(* Logix 5000 project; controller R400_500_XLS vendor 1 type 14 code 216 rev 31.11; software revision 31.01; part 23 of 32 *)
(* tags used below, declared in another part *)
   Abort1 : DINT;   // Not Used
   Alarm : SINT;   // Wait 3 seconds
   AlarmAcked : BOOL;   // Alarm has been acked
   bAlrm : BOOL[64];
   CycExcBuffer : UDT_CYCLE;
   CycleSequence : UDT_CYCLE_SEQUENCE;
   DrnSmp : DINT;
   DRYING : DINT;   // Drying id number
   drying_sp : REAL;   // Drying temperature set point
   drying_sp_offset : REAL;   // Low drying offset
   DRYING_TEMP_HIGH : REAL;   // Smart drying high temperature set point
   DRYING_TEMP_LOW : REAL;   // Smart drying low temperature set point
   DRYING_TEMP_STANDARD_LOW : REAL;   // Regular drying low temperature set point
   DRYING_TIME_LONG : DINT;   // Smart drying time for heat sensitive mode (in minute)
   DRYING_TIME_SHORT : DINT;   // Smart drying time for heat regular mode (in minute)
   dryingSmartTime : DINT;   // Duration of the smart drying phase
   DryingTempCool : REAL;   // Temperature limit for the smart drying mode cooling phase
   F2rinse : DINT;   // Not Used
   F3rinse : DINT;   // Not Used
   F4rinse : INT;   // Transition for the conductivity based evalutaion
   F4rinse_Tran : INT;   // Transitions for the conductivity based evaluation
   Fill_Sump : DINT;
   FRinseCondValue : REAL;   // Stored value of the conductivity
   HeatSmp : DINT;
   Inj_Time : SINT;   // Time based chemical injection steps
   M : DINT[5];   // Memory Bits
   NbFinalRinseDone : DINT;
   Neutral : SINT;
   ONS_FC08 : DINT;
   ONS_FC09 : SINT;
   PureWaterTankFilling : BOOL;   // Start PWT filling
   Run : DINT;
   STANDARD : SINT;
   SumpWaterVolume : DINT;   // Sump Water Volume 0 =Low 1= High
   Tmr : TIMER[107];
   Treatment_info : DINT;   // Treatment message conditions
   Trt_Drying : SINT;
   Trt_Drying_Tran : INT;
   Trt_Vapor_Exhaust : BOOL;   // Vapor exhaust fan is on
   VENTING : DINT;   // Venting id number
   WaterSaved : BOOL;   // Water Saved In Sump (Last Final Rinse Water)
   WSH56_TreatmentInfo : BOOL;   // Treatment information for the conductivity injection
   COOLING_PHASE_TIME : DINT;   // Time of the cooling phase when time based drying
   DryTemp : REAL;
   FALSE : BOOL;   // Always false bit
   FinalRinseCond : REAL;
   Msg_Phase : DINT;
   PrintFrinseCondValue : REAL;
   PureWaterTankDrainingDeadLeg : BOOL;
   PureWaterTankFillingRequest : BOOL;
   Q_Smp_Stm_Vlve : BOOL;   // Sump steam valve/ Electrical Heater
   TreatmentPtr : DINT;
   Unit : Hrdwre;   // Unit Configuration
(* MainProgram, continued *)

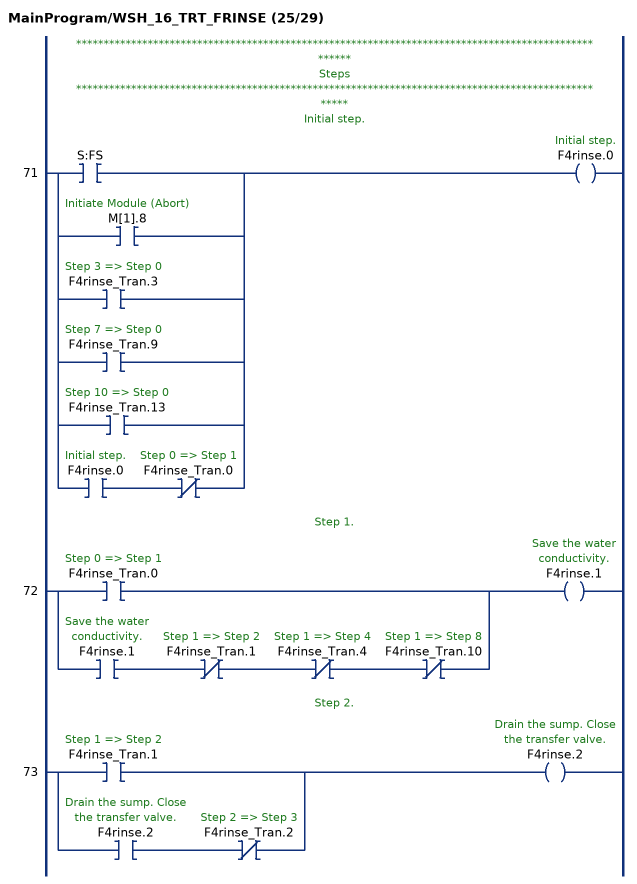
   [picture p449: MainProgram/WSH_16_TRT_FRINSE rungs 71-73]
   // ****************************************************************************************************
   // Steps
   // ***************************************************************************************************
   // Initial step.
   71: [XIC(S:FS) ,XIC(M[1].8) ,XIC(F4rinse_Tran.3) ,XIC(F4rinse_Tran.9) ,XIC(F4rinse_Tran.13) ,XIC(F4rinse.0) XIO(F4rinse_Tran.0) ]OTE(F4rinse.0);
   // Step 1.
   72: [XIC(F4rinse_Tran.0) ,XIC(F4rinse.1) XIO(F4rinse_Tran.1) XIO(F4rinse_Tran.4) XIO(F4rinse_Tran.10) ]OTE(F4rinse.1);
   // Step 2.
   73: [XIC(F4rinse_Tran.1) ,XIC(F4rinse.2) XIO(F4rinse_Tran.2) ]OTE(F4rinse.2);
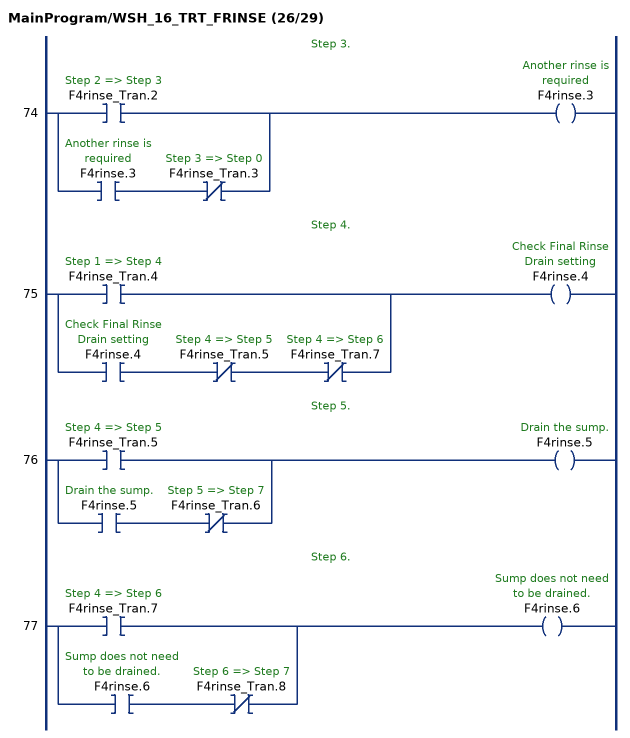
   // Step 3.
   74: [XIC(F4rinse_Tran.2) ,XIC(F4rinse.3) XIO(F4rinse_Tran.3) ]OTE(F4rinse.3);
   // Step 4.
   75: [XIC(F4rinse_Tran.4) ,XIC(F4rinse.4) XIO(F4rinse_Tran.5) XIO(F4rinse_Tran.7) ]OTE(F4rinse.4);
   // Step 5.
   76: [XIC(F4rinse_Tran.5) ,XIC(F4rinse.5) XIO(F4rinse_Tran.6) ]OTE(F4rinse.5);
   // Step 6.
   77: [XIC(F4rinse_Tran.7) ,XIC(F4rinse.6) XIO(F4rinse_Tran.8) ]OTE(F4rinse.6);
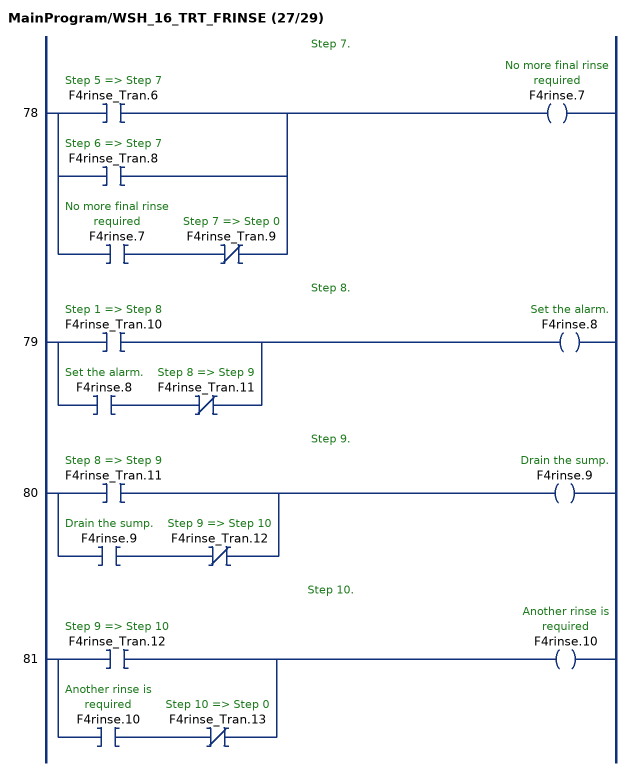
   // Step 7.
   78: [XIC(F4rinse_Tran.6) ,XIC(F4rinse_Tran.8) ,XIC(F4rinse.7) XIO(F4rinse_Tran.9) ]OTE(F4rinse.7);
   // Step 8.
   79: [XIC(F4rinse_Tran.10) ,XIC(F4rinse.8) XIO(F4rinse_Tran.11) ]OTE(F4rinse.8);
   // Step 9.
   80: [XIC(F4rinse_Tran.11) ,XIC(F4rinse.9) XIO(F4rinse_Tran.12) ]OTE(F4rinse.9);
   // Step 10.
   81: [XIC(F4rinse_Tran.12) ,XIC(F4rinse.10) XIO(F4rinse_Tran.13) ]OTE(F4rinse.10);
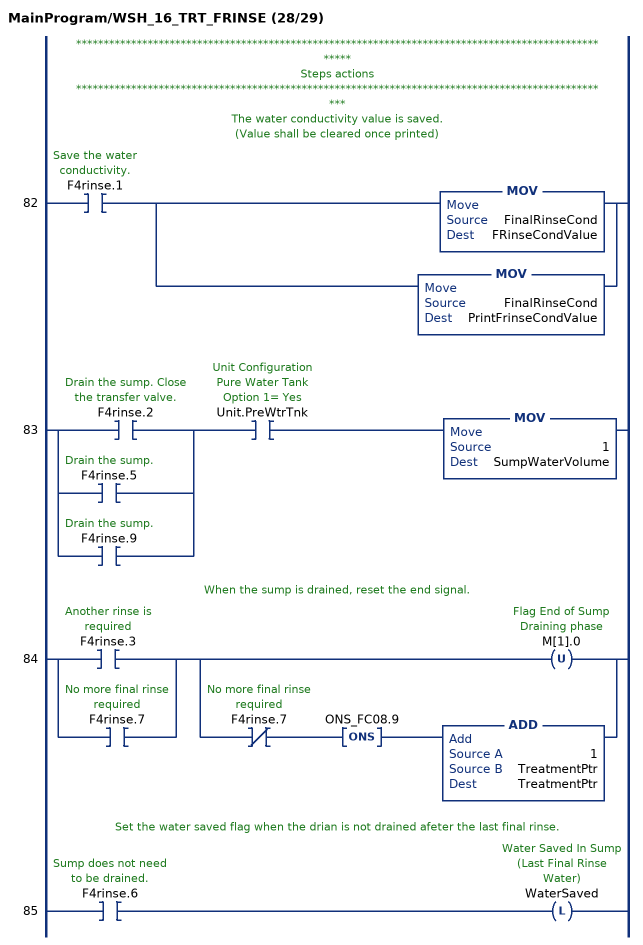
   // ****************************************************************************************************
   // Steps actions
   // **************************************************************************************************
   // The water conductivity value is saved.
   // (Value shall be cleared once printed)
   82: XIC(F4rinse.1)[MOV(FinalRinseCond,FRinseCondValue) ,MOV(FinalRinseCond,PrintFrinseCondValue) ];
   83: [XIC(F4rinse.2) ,XIC(F4rinse.5) ,XIC(F4rinse.9) ]XIC(Unit.PreWtrTnk)MOV(1,SumpWaterVolume);
   // When the sump is drained, reset the end signal.
   84: [XIC(F4rinse.3) ,XIC(F4rinse.7) ][OTU(M[1].0) ,XIO(F4rinse.7) ONS(ONS_FC08.9) ADD(1,TreatmentPtr,TreatmentPtr) ];
   // Set the water saved flag when the drian is not drained afeter the last final rinse.
   85: XIC(F4rinse.6)OTL(WaterSaved);
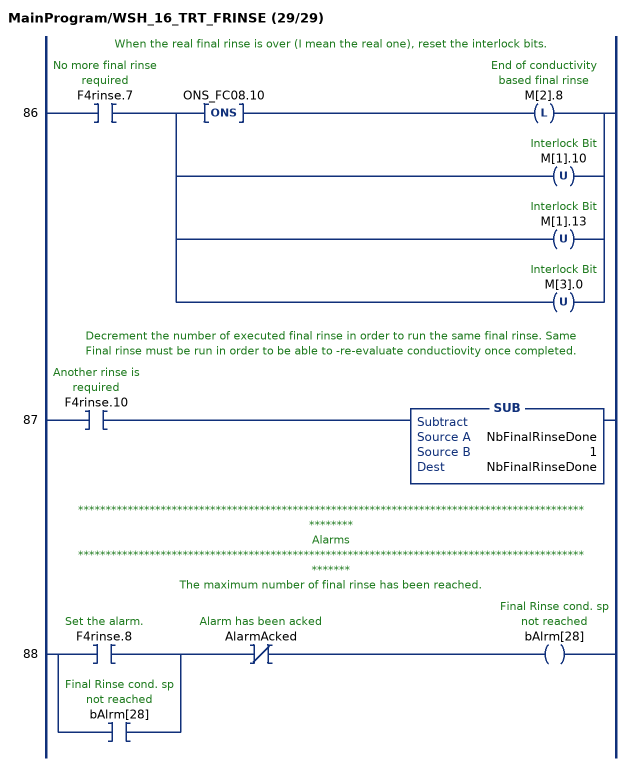
   // When the real final rinse is over (I mean the real one), reset the interlock bits.
   86: XIC(F4rinse.7)[ONS(ONS_FC08.10) OTL(M[2].8) ,OTU(M[1].10) ,OTU(M[1].13) ,OTU(M[3].0) ];
   // Decrement the number of executed final rinse in order to run the same final rinse. Same Final rinse must be run in order to be able to -re-evaluate conductiovity once completed.
   87: XIC(F4rinse.10)SUB(NbFinalRinseDone,1,NbFinalRinseDone);
   // ****************************************************************************************************
   // Alarms
   // ***************************************************************************************************
   // The maximum number of final rinse has been reached.
   88: [XIC(F4rinse.8) ,XIC(bAlrm[28]) ]XIO(AlarmAcked)OTE(bAlrm[28]);
END_ROUTINE

ROUTINE WSH_18_DRYING   (* ladder *)
// ROUTINe
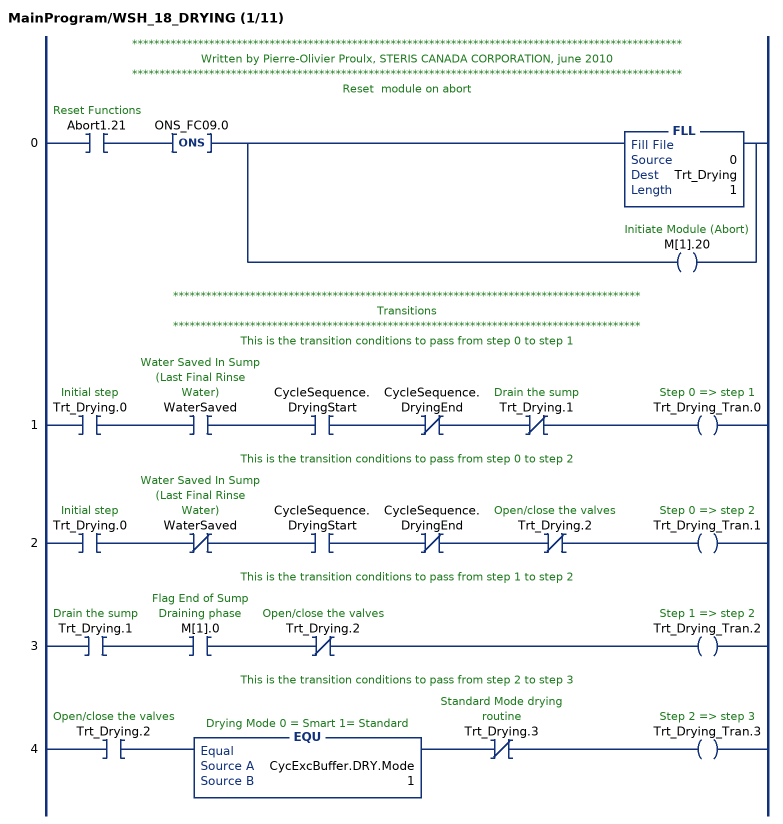
   // ****************************************************************************************************
   // Written by Pierre-Olivier Proulx, STERIS CANADA CORPORATION, june 2010
   // ****************************************************************************************************
   // Reset  module on abort
   0: XIC(Abort1.21)ONS(ONS_FC09.0)[FLL(0,Trt_Drying,1) ,OTE(M[1].20) ];
   // *************************************************************************************
   // Transitions
   // *************************************************************************************
   // This is the transition conditions to pass from step 0 to step 1
   1: XIC(Trt_Drying.0)XIC(WaterSaved)XIC(CycleSequence.DryingStart)XIO(CycleSequence.DryingEnd)XIO(Trt_Drying.1)OTE(Trt_Drying_Tran.0);
   // This is the transition conditions to pass from step 0 to step 2
   2: XIC(Trt_Drying.0)XIO(WaterSaved)XIC(CycleSequence.DryingStart)XIO(CycleSequence.DryingEnd)XIO(Trt_Drying.2)OTE(Trt_Drying_Tran.1);
   // This is the transition conditions to pass from step 1 to step 2
   3: XIC(Trt_Drying.1)XIC(M[1].0)XIO(Trt_Drying.2)OTE(Trt_Drying_Tran.2);
   // This is the transition conditions to pass from step 2 to step 3
   4: XIC(Trt_Drying.2)EQU(CycExcBuffer.DRY.Mode,1)XIO(Trt_Drying.3)OTE(Trt_Drying_Tran.3);
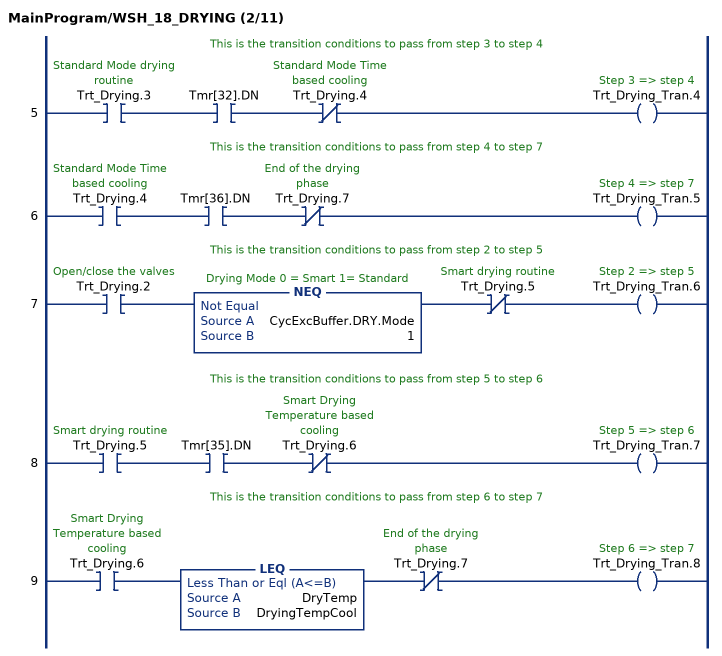
   // This is the transition conditions to pass from step 3 to step 4
   5: XIC(Trt_Drying.3)XIC(Tmr[32].DN)XIO(Trt_Drying.4)OTE(Trt_Drying_Tran.4);
   // This is the transition conditions to pass from step 4 to step 7
   6: XIC(Trt_Drying.4)XIC(Tmr[36].DN)XIO(Trt_Drying.7)OTE(Trt_Drying_Tran.5);
   // This is the transition conditions to pass from step 2 to step 5
   7: XIC(Trt_Drying.2)NEQ(CycExcBuffer.DRY.Mode,1)XIO(Trt_Drying.5)OTE(Trt_Drying_Tran.6);
   // This is the transition conditions to pass from step 5 to step 6
   8: XIC(Trt_Drying.5)XIC(Tmr[35].DN)XIO(Trt_Drying.6)OTE(Trt_Drying_Tran.7);
   // This is the transition conditions to pass from step 6 to step 7
   9: XIC(Trt_Drying.6)LEQ(DryTemp,DryingTempCool)XIO(Trt_Drying.7)OTE(Trt_Drying_Tran.8);
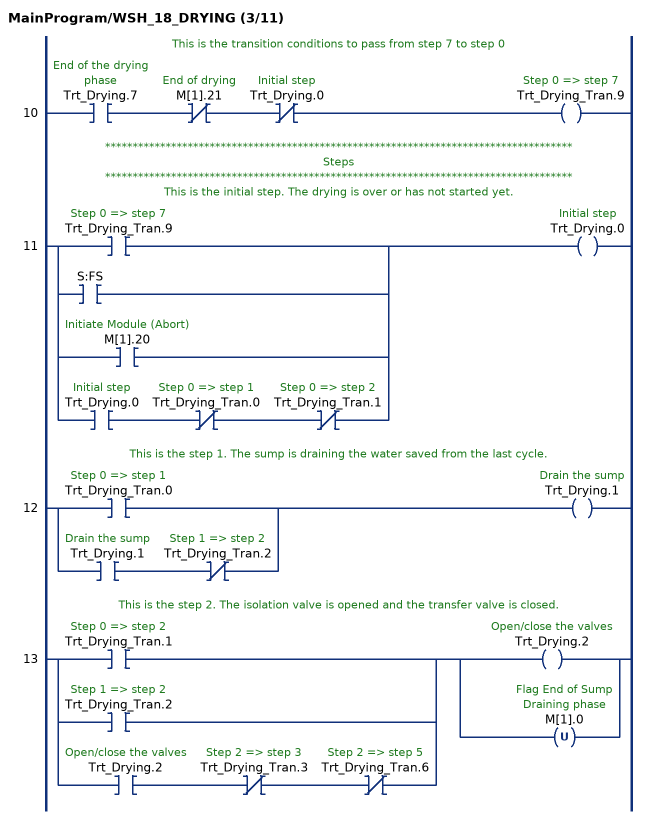
   // This is the transition conditions to pass from step 7 to step 0
   10: XIC(Trt_Drying.7)XIO(M[1].21)XIO(Trt_Drying.0)OTE(Trt_Drying_Tran.9);
   // *************************************************************************************
   // Steps
   // *************************************************************************************
   // This is the initial step. The drying is over or has not started yet.
   11: [XIC(Trt_Drying_Tran.9) ,XIC(S:FS) ,XIC(M[1].20) ,XIC(Trt_Drying.0) XIO(Trt_Drying_Tran.0) XIO(Trt_Drying_Tran.1) ]OTE(Trt_Drying.0);
   // This is the step 1. The sump is draining the water saved from the last cycle.
   12: [XIC(Trt_Drying_Tran.0) ,XIC(Trt_Drying.1) XIO(Trt_Drying_Tran.2) ]OTE(Trt_Drying.1);
   // This is the step 2. The isolation valve is opened and the transfer valve is closed.
   13: [XIC(Trt_Drying_Tran.1) ,XIC(Trt_Drying_Tran.2) ,XIC(Trt_Drying.2) XIO(Trt_Drying_Tran.3) XIO(Trt_Drying_Tran.6) ][OTE(Trt_Drying.2) ,OTU(M[1].0) ];
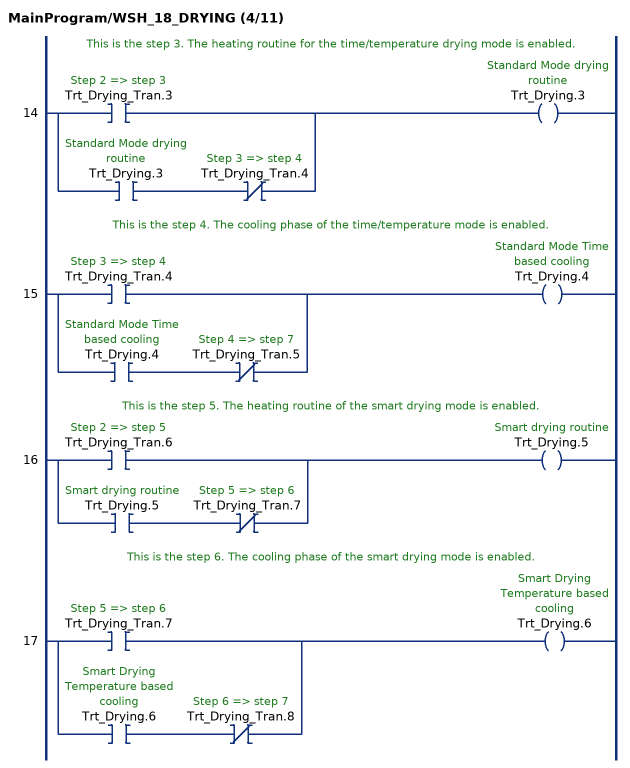
   // This is the step 3. The heating routine for the time/temperature drying mode is enabled.
   14: [XIC(Trt_Drying_Tran.3) ,XIC(Trt_Drying.3) XIO(Trt_Drying_Tran.4) ]OTE(Trt_Drying.3);
   // This is the step 4. The cooling phase of the time/temperature mode is enabled.
   15: [XIC(Trt_Drying_Tran.4) ,XIC(Trt_Drying.4) XIO(Trt_Drying_Tran.5) ]OTE(Trt_Drying.4);
   // This is the step 5. The heating routine of the smart drying mode is enabled.
   16: [XIC(Trt_Drying_Tran.6) ,XIC(Trt_Drying.5) XIO(Trt_Drying_Tran.7) ]OTE(Trt_Drying.5);
   // This is the step 6. The cooling phase of the smart drying mode is enabled.
   17: [XIC(Trt_Drying_Tran.7) ,XIC(Trt_Drying.6) XIO(Trt_Drying_Tran.8) ]OTE(Trt_Drying.6);
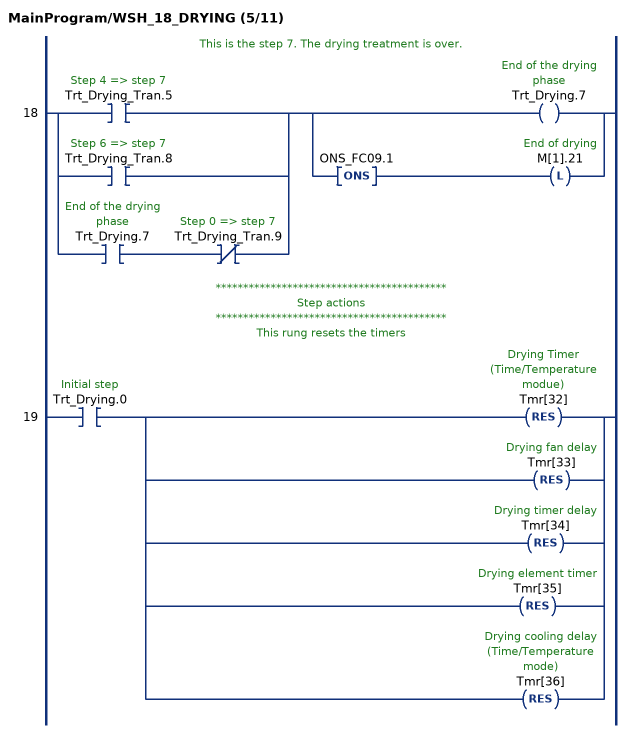
   // This is the step 7. The drying treatment is over.
   18: [XIC(Trt_Drying_Tran.5) ,XIC(Trt_Drying_Tran.8) ,XIC(Trt_Drying.7) XIO(Trt_Drying_Tran.9) ][OTE(Trt_Drying.7) ,ONS(ONS_FC09.1) OTL(M[1].21) ];
   // ******************************************
   // Step actions
   // ******************************************
   // This rung resets the timers
   19: XIC(Trt_Drying.0)[RES(Tmr[32]) ,RES(Tmr[33]) ,RES(Tmr[34]) ,RES(Tmr[35]) ,RES(Tmr[36]) ];
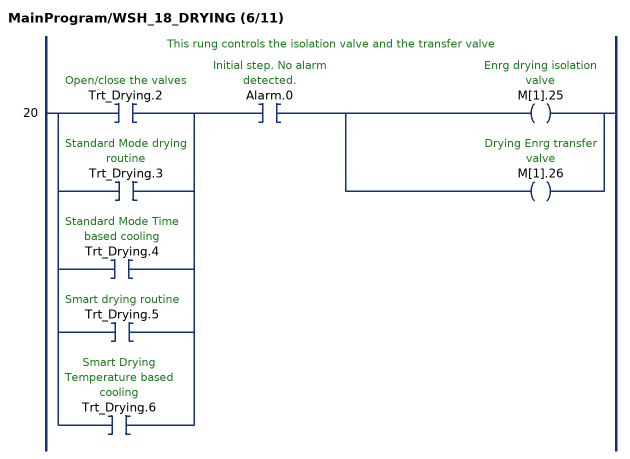
   // This rung controls the isolation valve and the transfer valve
   20: [XIC(Trt_Drying.2) ,XIC(Trt_Drying.3) ,XIC(Trt_Drying.4) ,XIC(Trt_Drying.5) ,XIC(Trt_Drying.6) ]XIC(Alarm.0)[OTE(M[1].25) ,OTE(M[1].26) ];
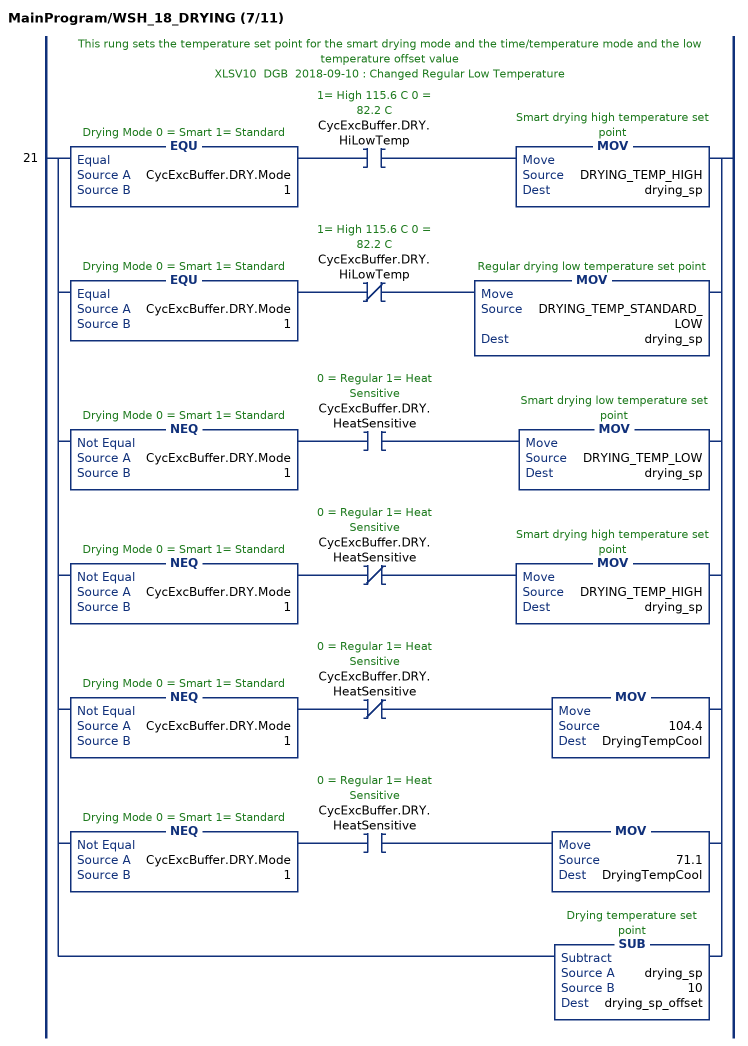
   // This rung sets the temperature set point for the smart drying mode and the time/temperature mode and the low temperature offset value
   // XLSV10  DGB  2018-09-10 : Changed Regular Low Temperature
   21: [EQU(CycExcBuffer.DRY.Mode,1) XIC(CycExcBuffer.DRY.HiLowTemp) MOV(DRYING_TEMP_HIGH,drying_sp) ,EQU(CycExcBuffer.DRY.Mode,1) XIO(CycExcBuffer.DRY.HiLowTemp) MOV(DRYING_TEMP_STANDARD_LOW,drying_sp) ,NEQ(CycExcBuffer.DRY.Mode,1) XIC(CycExcBuffer.DRY.HeatSensitive) MOV(DRYING_TEMP_LOW,drying_sp) ,NEQ(CycExcBuffer.DRY.Mode,1) XIO(CycExcBuffer.DRY.HeatSensitive) MOV(DRYING_TEMP_HIGH,drying_sp) ,NEQ(CycExcBuffer.DRY.Mode,1) XIO(CycExcBuffer.DRY.HeatSensitive) MOV(104.4,DryingTempCool) ,NEQ(CycExcBuffer.DRY.Mode,1) XIC(CycExcBuffer.DRY.HeatSensitive) MOV(71.1,DryingTempCool) ,SUB(drying_sp,10,drying_sp_offset) ];
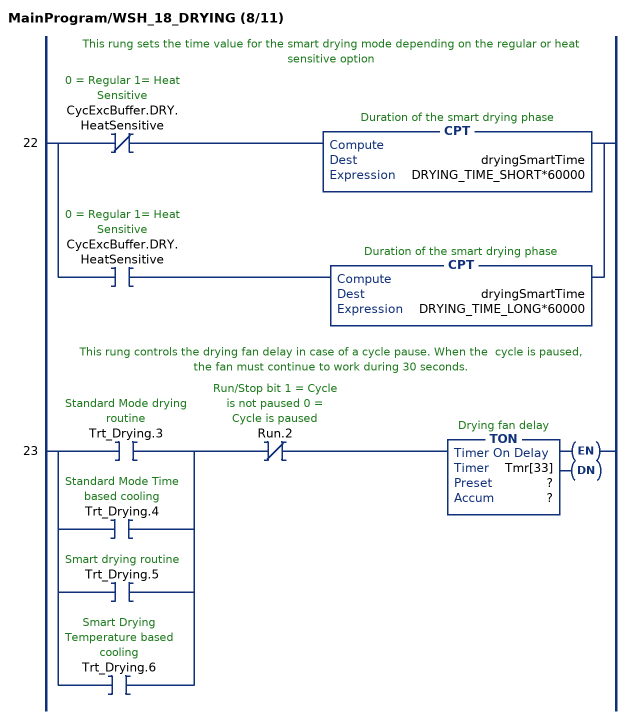
   // This rung sets the time value for the smart drying mode depending on the regular or heat sensitive option
   22: [XIO(CycExcBuffer.DRY.HeatSensitive) CPT(dryingSmartTime,DRYING_TIME_SHORT*60000) ,XIC(CycExcBuffer.DRY.HeatSensitive) CPT(dryingSmartTime,DRYING_TIME_LONG*60000) ];
   // This rung controls the drying fan delay in case of a cycle pause. When the  cycle is paused, the fan must continue to work during 30 seconds.
   23: [XIC(Trt_Drying.3) ,XIC(Trt_Drying.4) ,XIC(Trt_Drying.5) ,XIC(Trt_Drying.6) ]XIO(Run.2)TON(Tmr[33],?,?);
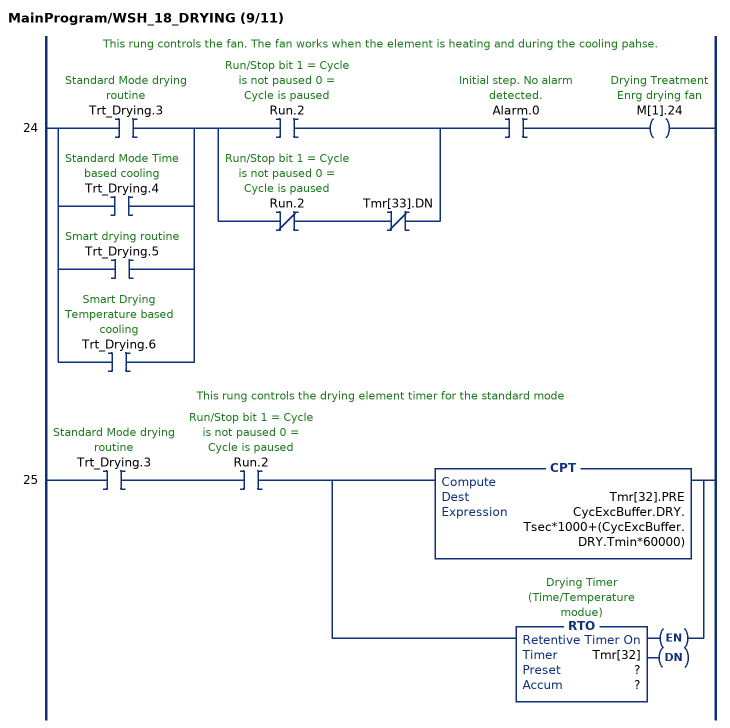
   // This rung controls the fan. The fan works when the element is heating and during the cooling pahse.
   24: [XIC(Trt_Drying.3) ,XIC(Trt_Drying.4) ,XIC(Trt_Drying.5) ,XIC(Trt_Drying.6) ][XIC(Run.2) ,XIO(Run.2) XIO(Tmr[33].DN) ]XIC(Alarm.0)OTE(M[1].24);
   // This rung controls the drying element timer for the standard mode
   25: XIC(Trt_Drying.3)XIC(Run.2)[CPT(Tmr[32].PRE,CycExcBuffer.DRY.Tsec*1000+(CycExcBuffer.DRY.Tmin*60000)) ,RTO(Tmr[32],?,?) ];
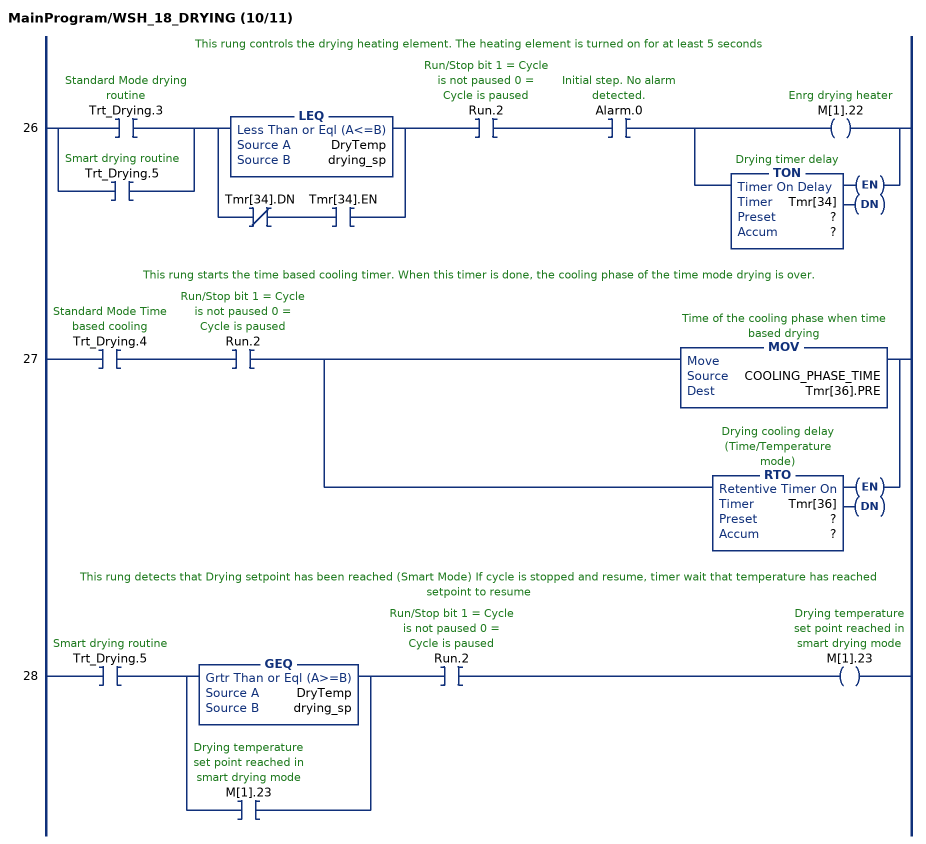
   // This rung controls the drying heating element. The heating element is turned on for at least 5 seconds
   26: [XIC(Trt_Drying.3) ,XIC(Trt_Drying.5) ][LEQ(DryTemp,drying_sp) ,XIO(Tmr[34].DN) XIC(Tmr[34].EN) ]XIC(Run.2)XIC(Alarm.0)[OTE(M[1].22) ,TON(Tmr[34],?,?) ];
   // This rung starts the time based cooling timer. When this timer is done, the cooling phase of the time mode drying is over.
   27: XIC(Trt_Drying.4)XIC(Run.2)[MOV(COOLING_PHASE_TIME,Tmr[36].PRE) ,RTO(Tmr[36],?,?) ];
   // This rung detects that Drying setpoint has been reached (Smart Mode) If cycle is stopped and resume, timer wait that temperature has reached setpoint to resume
   28: XIC(Trt_Drying.5)[GEQ(DryTemp,drying_sp) ,XIC(M[1].23) ]XIC(Run.2)OTE(M[1].23);
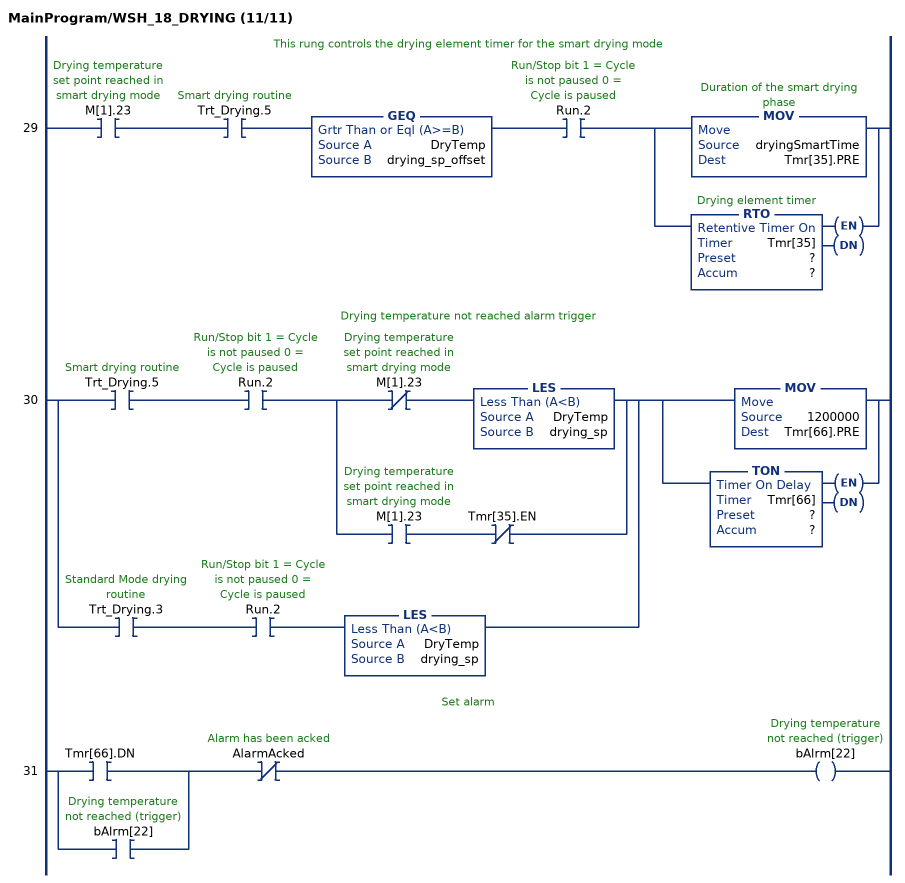
   // This rung controls the drying element timer for the smart drying mode
   29: XIC(M[1].23)XIC(Trt_Drying.5)GEQ(DryTemp,drying_sp_offset)XIC(Run.2)[MOV(dryingSmartTime,Tmr[35].PRE) ,RTO(Tmr[35],?,?) ];
   // Drying temperature not reached alarm trigger
   30: [XIC(Trt_Drying.5) XIC(Run.2) [XIO(M[1].23) LES(DryTemp,drying_sp) ,XIC(M[1].23) XIO(Tmr[35].EN) ] ,XIC(Trt_Drying.3) XIC(Run.2) LES(DryTemp,drying_sp) ][MOV(1200000,Tmr[66].PRE) ,TON(Tmr[66],?,?) ];
   // Set alarm
   31: [XIC(Tmr[66].DN) ,XIC(bAlrm[22]) ]XIO(AlarmAcked)OTE(bAlrm[22]);
END_ROUTINE

ROUTINE WSH_19_VENTING   (* ladder *)
// This routine vents the chamber
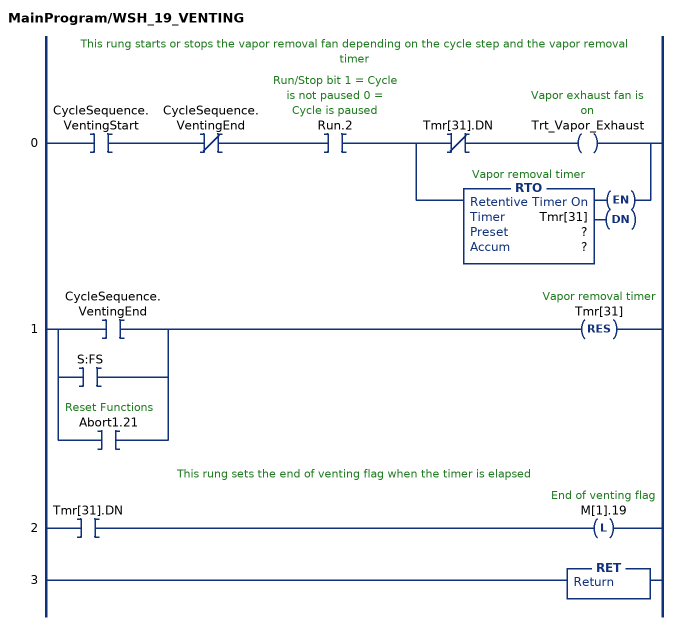
   // This rung starts or stops the vapor removal fan depending on the cycle step and the vapor removal timer
   0: XIC(CycleSequence.VentingStart)XIO(CycleSequence.VentingEnd)XIC(Run.2)[XIO(Tmr[31].DN) OTE(Trt_Vapor_Exhaust) ,RTO(Tmr[31],?,?) ];
   1: [XIC(CycleSequence.VentingEnd) ,[XIC(S:FS) ,XIC(Abort1.21) ] ]RES(Tmr[31]);
   // This rung sets the end of venting flag when the timer is elapsed
   2: XIC(Tmr[31].DN)OTL(M[1].19);
   3: RET();
END_ROUTINE

ROUTINE WSH_20_TREATMENT_INFO   (* ladder *)
// This routine decides which message the HMI will display during a cycle
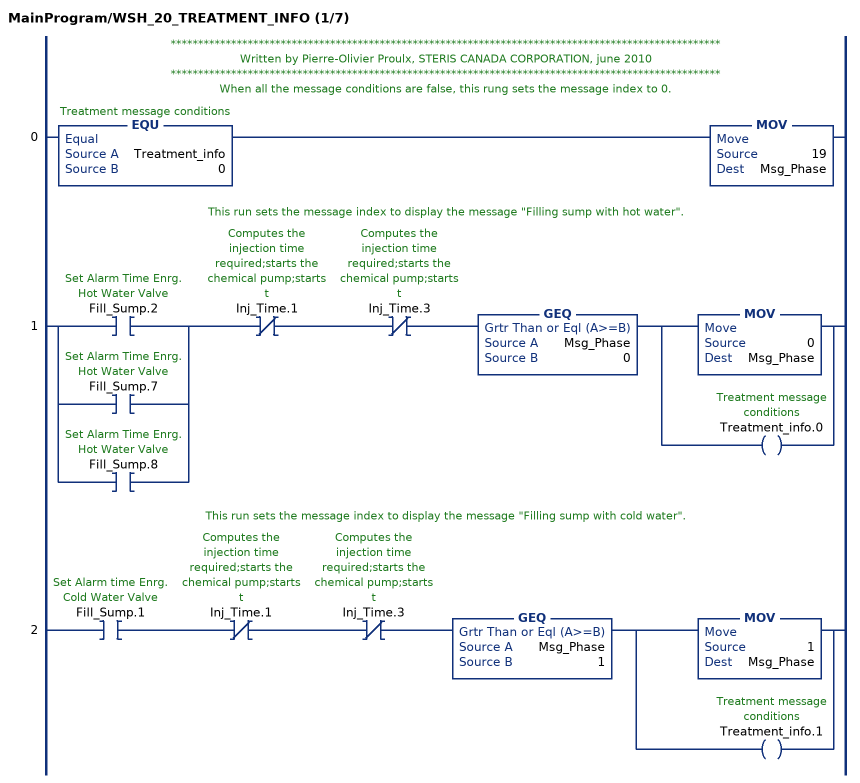
   // ****************************************************************************************************
   // Written by Pierre-Olivier Proulx, STERIS CANADA CORPORATION, june 2010
   // ****************************************************************************************************
   // When all the message conditions are false, this rung sets the message index to 0.
   0: EQU(Treatment_info,0)MOV(19,Msg_Phase);
   // This run sets the message index to display the message "Filling sump with hot water".
   1: [XIC(Fill_Sump.2) ,XIC(Fill_Sump.7) ,XIC(Fill_Sump.8) ]XIO(Inj_Time.1)XIO(Inj_Time.3)GEQ(Msg_Phase,0)[MOV(0,Msg_Phase) ,OTE(Treatment_info.0) ];
   // This run sets the message index to display the message "Filling sump with cold water".
   2: XIC(Fill_Sump.1)XIO(Inj_Time.1)XIO(Inj_Time.3)GEQ(Msg_Phase,1)[MOV(1,Msg_Phase) ,OTE(Treatment_info.1) ];
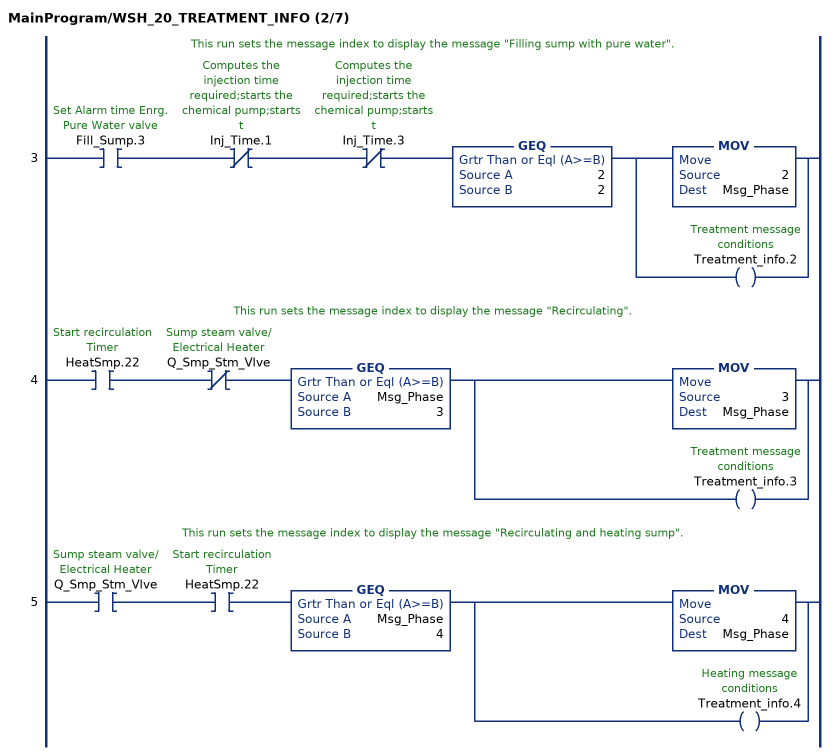
   // This run sets the message index to display the message "Filling sump with pure water".
   3: XIC(Fill_Sump.3)XIO(Inj_Time.1)XIO(Inj_Time.3)GEQ(2,2)[MOV(2,Msg_Phase) ,OTE(Treatment_info.2) ];
   // This run sets the message index to display the message "Recirculating".
   4: XIC(HeatSmp.22)XIO(Q_Smp_Stm_Vlve)GEQ(Msg_Phase,3)[MOV(3,Msg_Phase) ,OTE(Treatment_info.3) ];
   // This run sets the message index to display the message "Recirculating and heating sump".
   5: XIC(Q_Smp_Stm_Vlve)XIC(HeatSmp.22)GEQ(Msg_Phase,4)[MOV(4,Msg_Phase) ,OTE(Treatment_info.4) ];
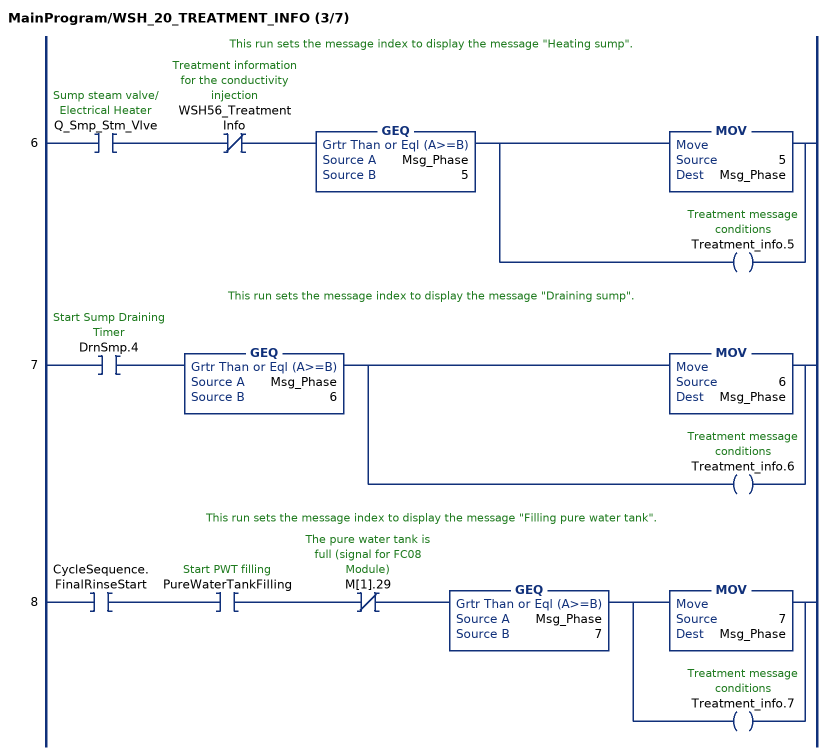
   // This run sets the message index to display the message "Heating sump".
   6: XIC(Q_Smp_Stm_Vlve)XIO(WSH56_TreatmentInfo)GEQ(Msg_Phase,5)[MOV(5,Msg_Phase) ,OTE(Treatment_info.5) ];
   // This run sets the message index to display the message "Draining sump".
   7: XIC(DrnSmp.4)GEQ(Msg_Phase,6)[MOV(6,Msg_Phase) ,OTE(Treatment_info.6) ];
   // This run sets the message index to display the message "Filling pure water tank".
   8: XIC(CycleSequence.FinalRinseStart)XIC(PureWaterTankFilling)XIO(M[1].29)GEQ(Msg_Phase,7)[MOV(7,Msg_Phase) ,OTE(Treatment_info.7) ];
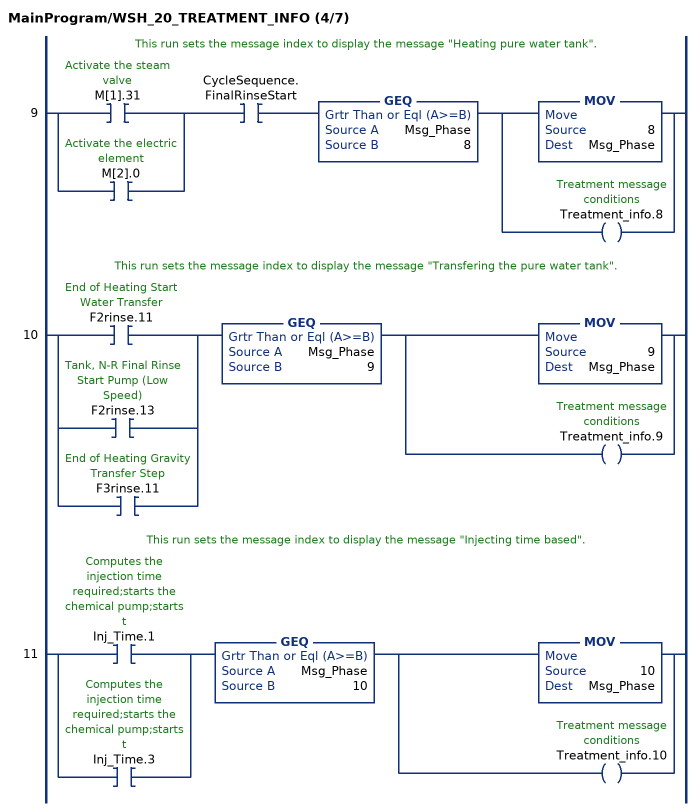
   // This run sets the message index to display the message "Heating pure water tank".
   9: [XIC(M[1].31) ,XIC(M[2].0) ]XIC(CycleSequence.FinalRinseStart)GEQ(Msg_Phase,8)[MOV(8,Msg_Phase) ,OTE(Treatment_info.8) ];
   // This run sets the message index to display the message "Transfering the pure water tank".
   10: [XIC(F2rinse.11) ,XIC(F2rinse.13) ,XIC(F3rinse.11) ]GEQ(Msg_Phase,9)[MOV(9,Msg_Phase) ,OTE(Treatment_info.9) ];
   // This run sets the message index to display the message "Injecting time based".
   11: [XIC(Inj_Time.1) ,XIC(Inj_Time.3) ]GEQ(Msg_Phase,10)[MOV(10,Msg_Phase) ,OTE(Treatment_info.10) ];
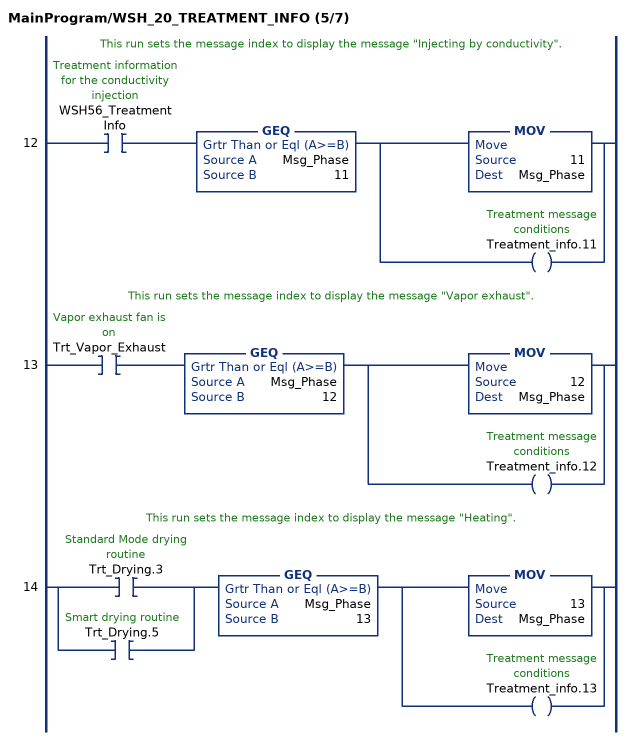
   // This run sets the message index to display the message "Injecting by conductivity".
   12: XIC(WSH56_TreatmentInfo)GEQ(Msg_Phase,11)[MOV(11,Msg_Phase) ,OTE(Treatment_info.11) ];
   // This run sets the message index to display the message "Vapor exhaust".
   13: XIC(Trt_Vapor_Exhaust)GEQ(Msg_Phase,12)[MOV(12,Msg_Phase) ,OTE(Treatment_info.12) ];
   // This run sets the message index to display the message "Heating".
   14: [XIC(Trt_Drying.3) ,XIC(Trt_Drying.5) ]GEQ(Msg_Phase,13)[MOV(13,Msg_Phase) ,OTE(Treatment_info.13) ];
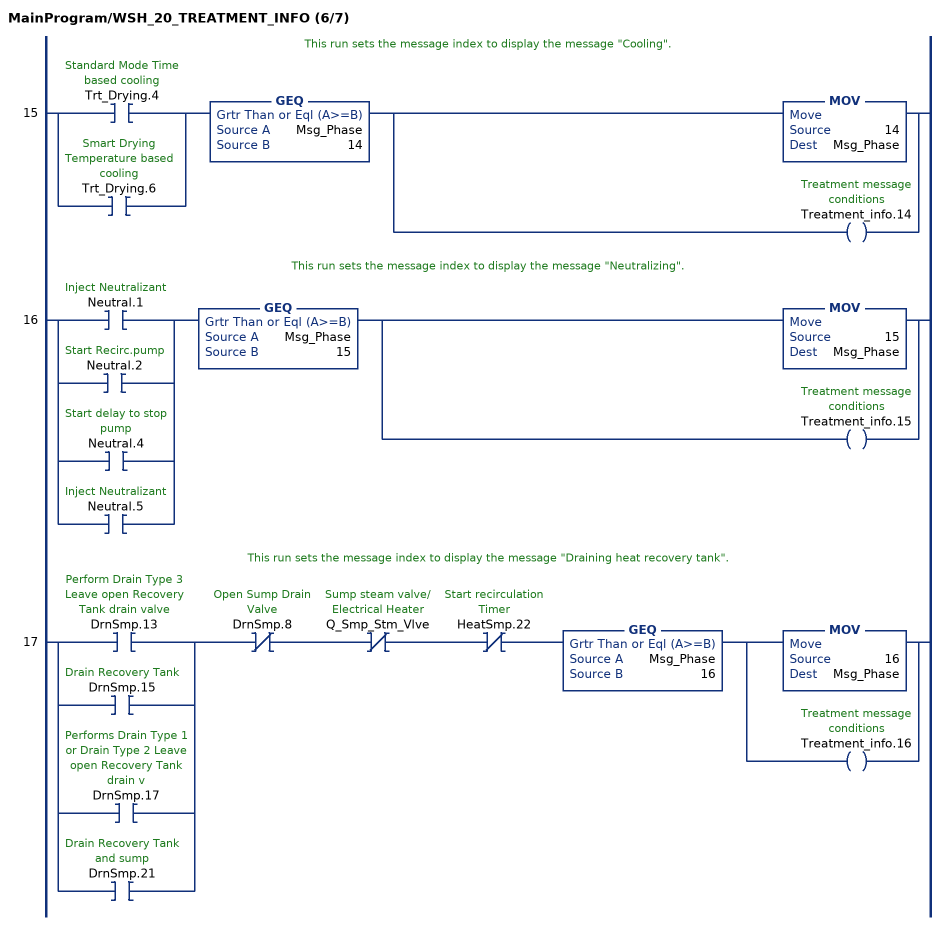
   // This run sets the message index to display the message "Cooling".
   15: [XIC(Trt_Drying.4) ,XIC(Trt_Drying.6) ]GEQ(Msg_Phase,14)[MOV(14,Msg_Phase) ,OTE(Treatment_info.14) ];
   // This run sets the message index to display the message "Neutralizing".
   16: [XIC(Neutral.1) ,XIC(Neutral.2) ,XIC(Neutral.4) ,XIC(Neutral.5) ]GEQ(Msg_Phase,15)[MOV(15,Msg_Phase) ,OTE(Treatment_info.15) ];
   // This run sets the message index to display the message "Draining heat recovery tank".
   17: [XIC(DrnSmp.13) ,XIC(DrnSmp.15) ,XIC(DrnSmp.17) ,XIC(DrnSmp.21) ]XIO(DrnSmp.8)XIO(Q_Smp_Stm_Vlve)XIO(HeatSmp.22)GEQ(Msg_Phase,16)[MOV(16,Msg_Phase) ,OTE(Treatment_info.16) ];
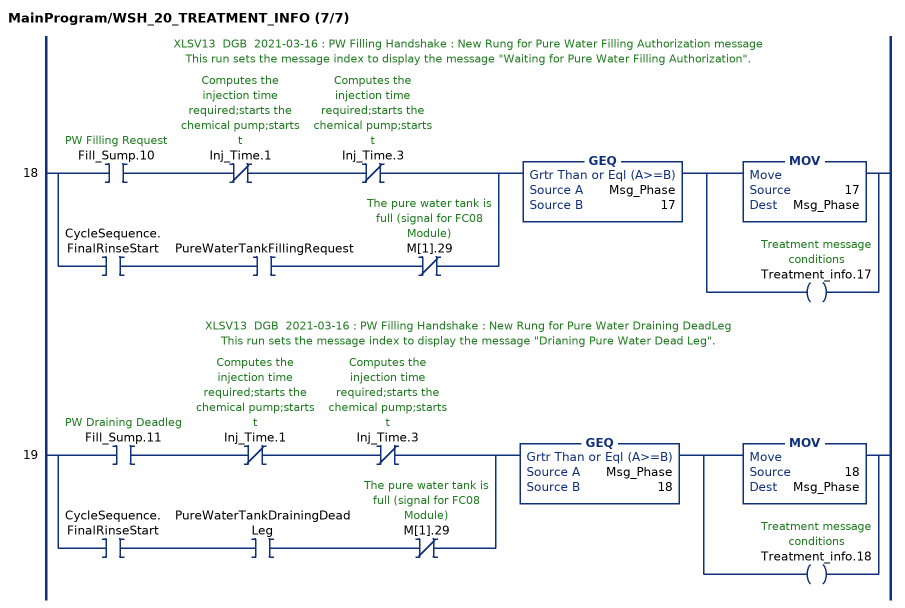
   // XLSV13  DGB  2021-03-16 : PW Filling Handshake : New Rung for Pure Water Filling Authorization message
   // This run sets the message index to display the message "Waiting for Pure Water Filling Authorization".
   18: [XIC(Fill_Sump.10) XIO(Inj_Time.1) XIO(Inj_Time.3) ,XIC(CycleSequence.FinalRinseStart) XIC(PureWaterTankFillingRequest) XIO(M[1].29) ]GEQ(Msg_Phase,17)[MOV(17,Msg_Phase) ,OTE(Treatment_info.17) ];
   // XLSV13  DGB  2021-03-16 : PW Filling Handshake : New Rung for Pure Water Draining DeadLeg
   // This run sets the message index to display the message "Drianing Pure Water Dead Leg".
   19: [XIC(Fill_Sump.11) XIO(Inj_Time.1) XIO(Inj_Time.3) ,XIC(CycleSequence.FinalRinseStart) XIC(PureWaterTankDrainingDeadLeg) XIO(M[1].29) ]GEQ(Msg_Phase,18)[MOV(18,Msg_Phase) ,OTE(Treatment_info.18) ];
END_ROUTINE
